PROGRAM main
  VAR
    S1 AT %IX0.0  : BOOL; (* botón del peatón *)
    SA1 AT %IX0.1 : BOOL; (* modo noche *)
    H1 AT %QX0.0  : BOOL; (* rojo *)
    H2 AT %QX0.1  : BOOL; (* amarillo *)
    H3 AT %QX0.2  : BOOL; (* verde *)
    H4 AT %QX0.3  : BOOL; (* verde peatonal *)
    X1            : BOOL; (* etapa VERDE *)
    X2            : BOOL; (* etapa AMARILLO *)
    X3            : BOOL; (* etapa ROJO *)
    T1            : BOOL; (* transición VERDE → AMARILLO *)
    T2            : BOOL; (* transición AMARILLO → ROJO *)
    T3            : BOOL; (* transición ROJO → VERDE *)
    ARRANQUE      : BOOL; (* solo en la primera vuelta *)
    INICIADO      : BOOL;
    PEATON        : BOOL; (* pedido del peatón *)
    PIDE          : BOOL; (* peatón o verde máximo *)
    T_VMIN        : TON;
    T_VMAX        : TON;
    T_AMA         : TON;
    T_ROJO        : TON;
    FIN_VMIN      : BOOL;
    FIN_VMAX      : BOOL;
    FIN_AMA       : BOOL;
    FIN_ROJO      : BOOL;
    T_ULT         : TON;
    ULTIMOS       : BOOL; (* últimos 3 s del rojo *)
    T_ON          : TON;
    T_OFF         : TON;
    ENCENDIDO     : BOOL;
    APAGADO       : BOOL;
    AMA_NORMAL    : BOOL;
  END_VAR
  VAR  (* added by the conversion: wires and edge detectors of the diagram *)
    _NOT1_OUT : BOOL;
    _OR4_OUT : BOOL;
    _OR24_OUT : BOOL;
    _AND28_OUT : BOOL;
    _AND33_OUT : BOOL;
    _AND37_OUT : BOOL;
    _OR42_OUT : BOOL;
    _NOT46_OUT : BOOL;
    _AND41_OUT : BOOL;
    _OR50_OUT : BOOL;
    _NOT53_OUT : BOOL;
    _AND49_OUT : BOOL;
    _OR57_OUT : BOOL;
    _NOT60_OUT : BOOL;
    _AND56_OUT : BOOL;
    _OR64_OUT : BOOL;
    _NOT67_OUT : BOOL;
    _AND63_OUT : BOOL;
  END_VAR

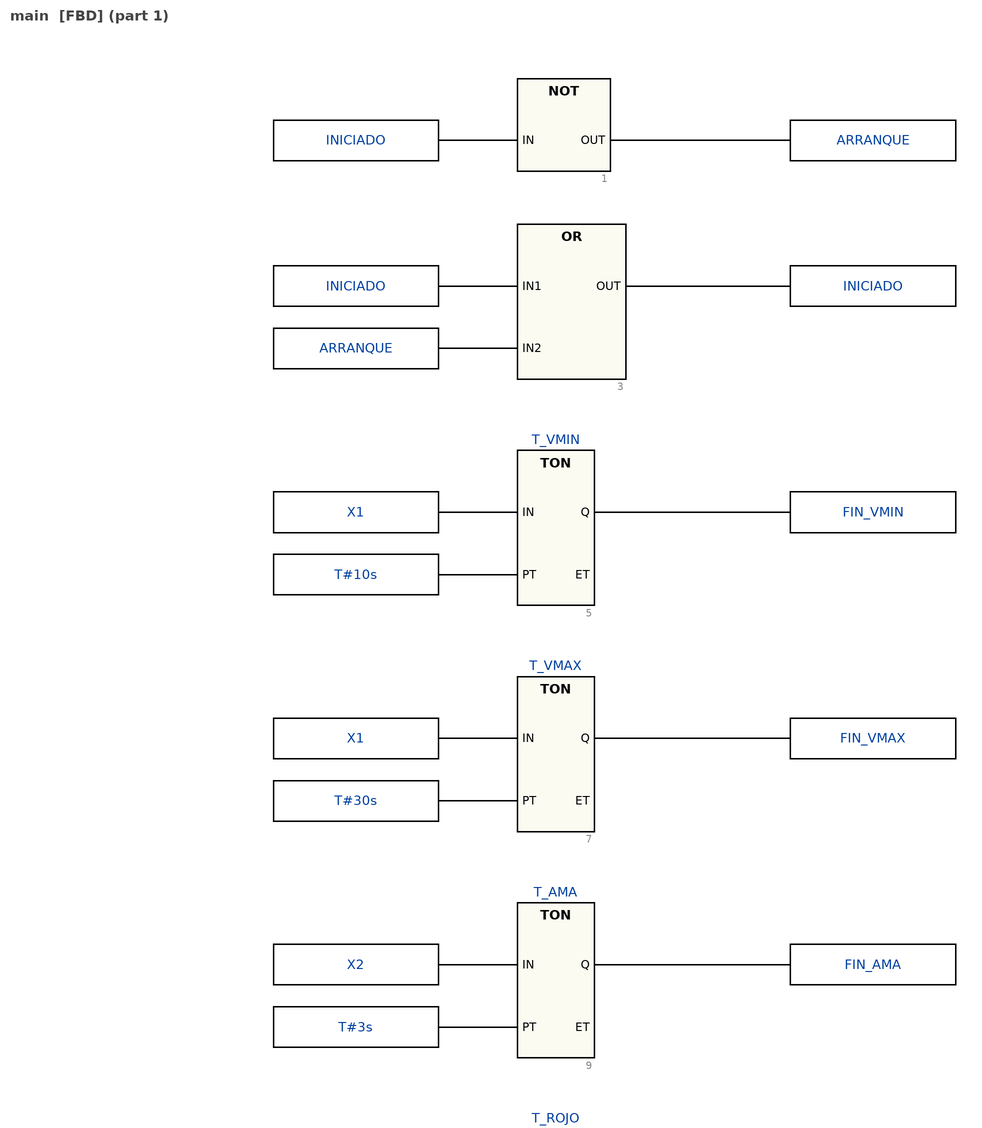
(* FBD diagram, written out as Structured Text *)
_NOT1_OUT := NOT INICIADO;
ARRANQUE := _NOT1_OUT;
_OR4_OUT := INICIADO OR ARRANQUE;
INICIADO := _OR4_OUT;
T_VMIN(IN := X1, PT := T#10s);
FIN_VMIN := T_VMIN.Q;
T_VMAX(IN := X1, PT := T#30s);
FIN_VMAX := T_VMAX.Q;
T_AMA(IN := X2, PT := T#3s);
FIN_AMA := T_AMA.Q;
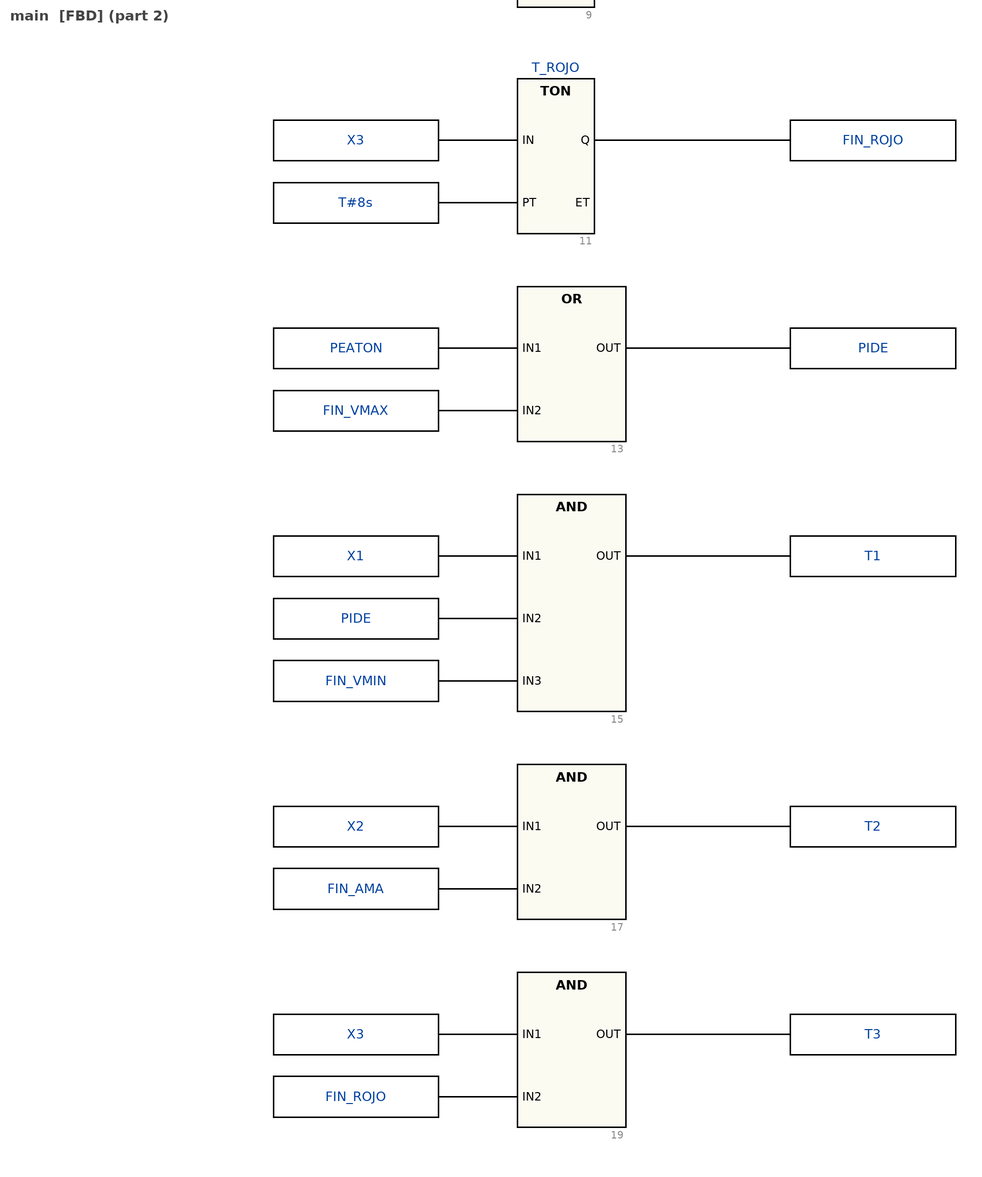
T_ROJO(IN := X3, PT := T#8s);
FIN_ROJO := T_ROJO.Q;
_OR24_OUT := PEATON OR FIN_VMAX;
PIDE := _OR24_OUT;
_AND28_OUT := X1 AND PIDE AND FIN_VMIN;
T1 := _AND28_OUT;
_AND33_OUT := X2 AND FIN_AMA;
T2 := _AND33_OUT;
_AND37_OUT := X3 AND FIN_ROJO;
T3 := _AND37_OUT;
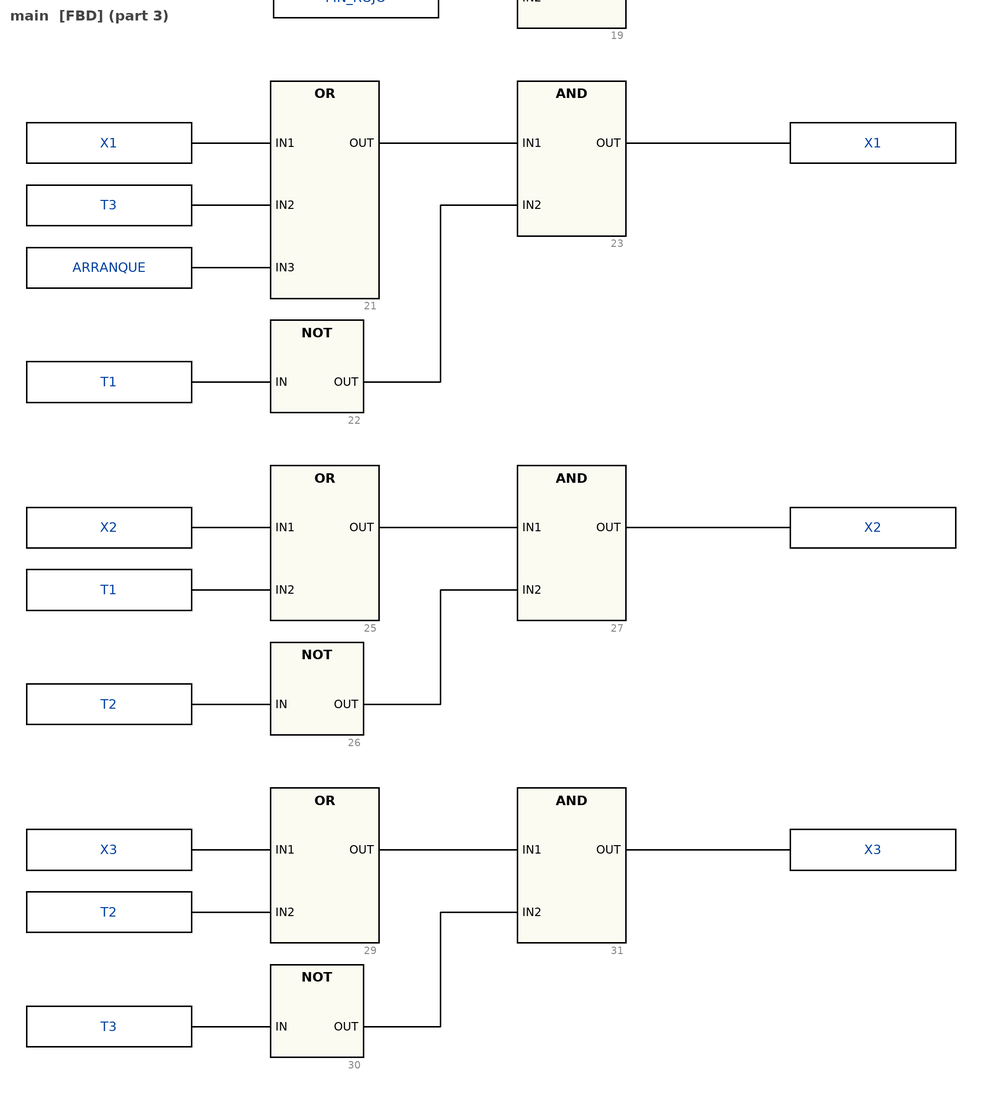
_OR42_OUT := X1 OR T3 OR ARRANQUE;
_NOT46_OUT := NOT T1;
_AND41_OUT := _OR42_OUT AND _NOT46_OUT;
X1 := _AND41_OUT;
_OR50_OUT := X2 OR T1;
_NOT53_OUT := NOT T2;
_AND49_OUT := _OR50_OUT AND _NOT53_OUT;
X2 := _AND49_OUT;
_OR57_OUT := X3 OR T2;
_NOT60_OUT := NOT T3;
_AND56_OUT := _OR57_OUT AND _NOT60_OUT;
X3 := _AND56_OUT;
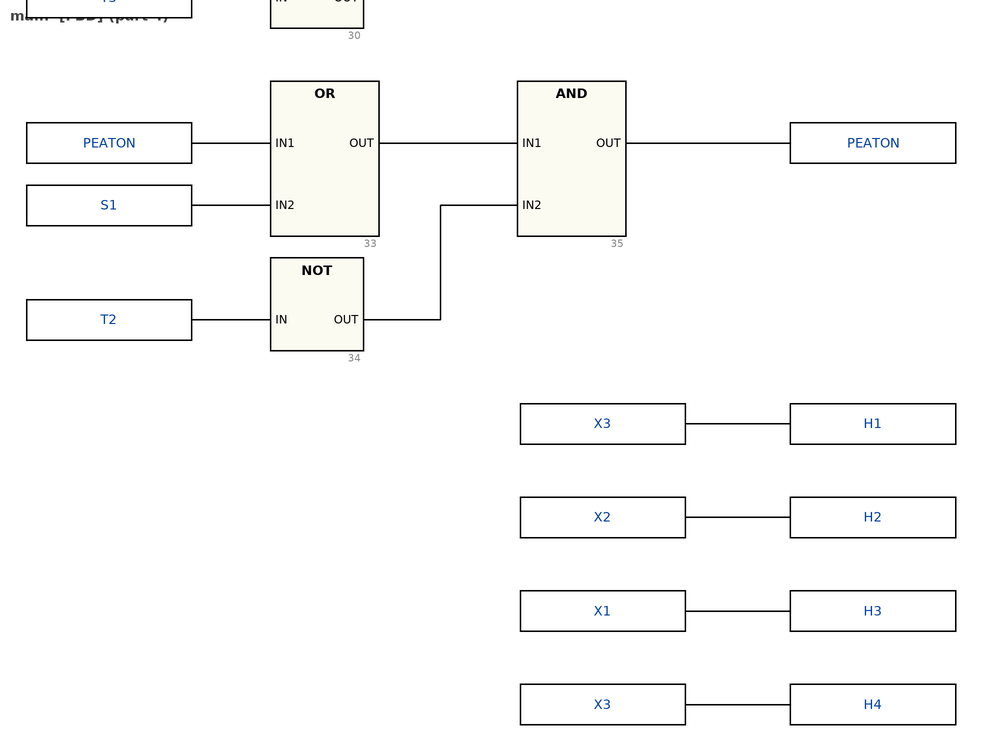
_OR64_OUT := PEATON OR S1;
_NOT67_OUT := NOT T2;
_AND63_OUT := _OR64_OUT AND _NOT67_OUT;
PEATON := _AND63_OUT;
H1 := X3;
H2 := X2;
H3 := X1;
H4 := X3;
END_PROGRAM
